(* IEC 61131-3 sources: NachHouse_TST/OSCAT_BasicLib/OscatBasicLib_333a, 28 files *)

(* ---- Arrays.ST ---- *)
TYPE
  OSCAT_BASIC_ARRAY0_32000_OF_REAL : ARRAY[0..32000] OF REAL;
  OSCAT_BASIC_ARRAY1_32000_OF_REAL : ARRAY[1..32000] OF REAL;
END_TYPE

(* @PATH := '\/Mathematical\/Array' *)
FUNCTION _ARRAY_ABS : BOOL
(*
  this function will calculate the absolute value of each element of the array and stroe the result instead of the element.
  Array[i] := ABS(ARRAY[i]).
  the function needs to be called:  array_avg(adr("array"),sizeof("array"));
  because this function works with pointers its very time efficient and it needs no extra memory.

  version 1.0 2. apr. 2008
  programmer  hugo
  tested by tobias
*)
  VAR_INPUT
    pt : PTR_TO OSCAT_BASIC_ARRAY0_32000_OF_REAL;
    size : UINT;
  END_VAR
  VAR
    i: UINT;
    stop: UINT;
  END_VAR

  stop := WORD_TO_UINT(SHR(UINT_TO_WORD(size),2))-1;
  FOR i := 0 TO stop DO
    PT^[i] := ABS(PT^[i]);
  END_FOR;
  _ARRAY_ABS := TRUE;

(* revision history
  hm  2. apr 2008   rev 1.0
    original version
*)
END_FUNCTION

(* @PATH := '\/Mathematical\/Array' *)
FUNCTION _ARRAY_ADD : BOOL
(*
  this function will add an offset X to each element of the array and stroe the result instead of the element.
  Array[i] := ARRAY[i] + X.
  the function needs to be called:  array_avg(adr("array"),sizeof("array"));
  because this function works with pointers its very time efficient and it needs no extra memory.

  version 1.0 2. apr. 2008
  programmer  hugo
  tested by tobias
*)
  VAR_INPUT
    pt : PTR_TO OSCAT_BASIC_ARRAY0_32000_OF_REAL;
    size : UINT;
    X : REAL;
  END_VAR
  VAR
    i: UINT;
    stop: UINT;
  END_VAR

  stop := WORD_TO_UINT(SHR(UINT_TO_WORD(size),2))-1; //SHR(size,2)-1;
  FOR i := 0 TO stop DO
    PT^[i] := PT^[i] + X;
  END_FOR;
  _ARRAY_ADD := TRUE;

(* revision history
  hm  2. apr 2008   rev 1.0
    original version
*)
END_FUNCTION

(* @PATH := '\/Mathematical\/Array' *)
FUNCTION _ARRAY_INIT : BOOL
(*
  this function will initialize a given array with a value init.
  the function needs to be called:  _array_init(adr("array"),sizeof("array"));
  this function will manipulate a given array.
  the function manipulates the original array, it rerturnes true when finished.
  because this function works with pointers its very time efficient and it needs no extra memory.

  version 1.3 16 mar 2008
  programmer  hugo
  tested by   tobias
*)
  VAR_INPUT
    pt : PTR_TO OSCAT_BASIC_ARRAY0_32000_OF_REAL;
    size : UINT;
    init : REAL;
  END_VAR
  VAR
    i: UINT;
    stop: UINT;
  END_VAR

  stop := WORD_TO_UINT(SHR(UINT_TO_WORD(size),2))-1; //SHR(size,2)-1;
  FOR i := 0 TO stop DO
    pt^[i] := init;
  END_FOR;

  _array_init := TRUE;

(* revision History
  hm 6.1.2007   rev 1.1
    change type of function to bool
    added  array_init := true to set output true.

  hm  14.11.2007  rev 1.2
    changed stop calculation to be more efficient

  hm  16.3. 2008    rev 1.3
    changed type of input size to uint
*)
END_FUNCTION

(* @PATH := '\/Mathematical\/Array' *)
FUNCTION _ARRAY_SORT : BOOL
(*
  this function will sort a given array.
  the function needs to be called:  _array_sort(adr("array"),sizeof("array"));
  this function will manipulate a given array.
  the function will not return anything except true, it will instead manipulate the original array.
  because this function works with pointers its very time efficient and it needs no extra memory.

  version 2.0 19. jan. 2011
  programmer  Alexander Trikitis
  tested by oscat
*)
  VAR_INPUT
    PT : PTR_TO OSCAT_BASIC_ARRAY1_32000_OF_REAL; // ARRAY[1..32000] OF REAL;
    SIZE : UINT;
  END_VAR
  VAR
    stack_count: UINT;        (* Laufvariable Stack*)
    stack: ARRAY[1..32] OF UINT;  (* Stackgröße~ 1,6*Log(n)/log(2) *)
                      (* Stackgröße 32 => ~1 Mio Elemente *)
    links: UINT;            (* Anfangselement des Arrays *)
    rechts: UINT;           (* Endelement des Arrays *)
    pivot: REAL;            (* temporärer Schwellwert für Tauschbedingung *)
    i: UINT;              (* Laufvariable1 *)
    j: UINT;              (* Laufvariable2 *)
    ende_innen: BOOL;       (* Ende innere Schleife *)
    ende_aussen: BOOL;        (* Ende äußere Schleife *)
    tmp: REAL;            (* Hilfsvariable zum Tauschen von Werten *)
  END_VAR

  (* Startwerte zur Arraygröße *)
  links := 1;         (* Anfangselement des Arrays *)
  rechts :=  WORD_TO_UINT(SHR(UINT_TO_WORD(size),2)); //SHR(size,2);    (* Endelement des Arrays *)
  stack_count := 1;     (* Laufvariable Stack *)

  WHILE NOT ende_aussen DO            (* äußere Schleife *)
    IF links < rechts THEN
      pivot := PT^[WORD_TO_UINT(SHR(UINT_TO_WORD(rechts+links),1))];      (* Wert des mittleren Elements als Pivot-Wert *)
      i := links -1;
      j := rechts +1;

      (* innere Schleife, teile Feld *)
      ende_innen := FALSE;
      REPEAT

        (* steigende Reihenfolge *)
        REPEAT  i := i+1; UNTIL (PT^[i] >= pivot) OR NOT (i < rechts) END_REPEAT;
        REPEAT  j := j-1; UNTIL (PT^[j] <= pivot) OR NOT (j > links)  END_REPEAT;

        (*sinkende Reihenfolge *)
  (*      REPEAT  i := i+1; UNTIL (PT^[i] <= pivot) OR NOT (i < rechts) END_REPEAT  *)
  (*      REPEAT  j := j-1; UNTIL (PT^[j] >= pivot) OR NOT (j > links)  END_REPEAT  *)

        IF i >= j THEN
          ende_innen := TRUE;
        ELSE
             tmp := PT^[j];
          PT^[j] := PT^[i];
          PT^[i] := tmp;
        END_IF;

      UNTIL ende_innen END_REPEAT;

      (* Push stack *)
      stack[stack_count] := rechts;   (* rechten Teil später sortieren *)
      IF Stack_count < 32 THEN
        stack_count := stack_count +1;
      ELSE
        ende_aussen := TRUE;
        _ARRAY_SORT := FALSE;         (* Fehler: Stack zu klein *)
      END_IF;

      (* linken Teil sortiern *)
      rechts := MAX(links, i-1);

    ELSE

      IF stack_count = 1 THEN
        ende_aussen := TRUE;
      ELSE

        links := rechts+1;

        (* pop stack *)
        stack_count := stack_count -1;    (* jetzt rechten Teil sortierne *)
        rechts:= stack[stack_count];
      END_IF;

    END_IF;

  END_WHILE;

  _ARRAY_SORT := TRUE;        (* Sortierung beendet *)

(* algorithm used before rev 2.0
  size := SHR(size,2);
  size2 := UINT_TO_INT(SHR(size,1));
  FOR i := SIZE2  TO 1 BY -1 DO
    j:=i;
      WHILE j <= SIZE2 DO
        stop := j * 2 + 1;
          IF stop > UINT_TO_INT(SIZE) THEN stop := stop - 1;
          ELSIF pt^[stop-1] > pt^[stop] THEN stop := stop - 1;
      END_IF;
          IF pt^[j] < pt^[stop] THEN
            temp := pt^[j];
              pt^[j] := pt^[stop];
              pt^[stop] := temp;
          END_IF;
          j := stop;
      END_WHILE;
  END_FOR;
*)

(* heapsort
  FOR heapsize := UINT_TO_INT(size) TO 1 BY -1 DO
    popmax := pt^[1];
    pt^[1] := pt^[heapsize];
      i := 1;
    hs2 := SHR(heapsize,1);
    WHILE i <= hs2 DO
          stop := i * 2 + 1;
            IF stop > heapsize THEN stop := stop - 1;
            ELSIF pt^[stop-1] > pt^[stop] THEN stop := stop - 1;
      END_IF;
            IF pt^[i] < pt^[stop] THEN
                  temp := pt^[i];
                  pt^[i] := pt^[stop];
                  pt^[stop] := temp;
            END_IF;
            i := stop;
        END_WHILE;
    pt^[heapsize] := popmax;
  END_FOR;

  _ARRAY_SORT2 := TRUE;
*)

(* old algorithm bubble sort used before rev 1.2
  stop := (size - SIZEOF(pt)) / SIZEOF(pt);
  FOR i := 0 TO stop - 1 DO
    FOR m := i + 1 TO stop DO
      IF pt^[i] > pt^[m] THEN
        temp := pt^[i];
        pt^[i] := pt^[m];
        pt^[m] := temp;
      END_IF;
    END_FOR;
  END_FOR;
  _array_sort := TRUE;
*)

(* revision history
  hm  6.1.2007  rev 1.1
    changed return value to true

  hm  22. sep 2007  rev 1.2
    changed sorting algorithm to heap sort for performance reasons

  hm  14. nov 2007  rev 1.3
    changed calculation of stop to be more efficient

  hm  15 dec 2007 rev 1.4
    added function return true

  hm  5. jan 2008   rev 1.5
    improved performance

  hm  16. mar. 2008 rev 1.6
    changed type of input size to uint

  hm  28. mar. 2008 rev 1.7
    changed input f to pt

  hm  19. jan. 2011 rev 2.0
    new faster algorithm using qucksort (Alexander Drikitis)
*)
END_FUNCTION

(* @PATH := '\/Mathematical\/Array' *)
FUNCTION _ARRAY_MEDIAN : REAL
(*
  this function will calculate the median of a given array.
  in order to do so the ariginal array is sorted and stays sorted after the function finishes
  the function needs to be called:  _array_median(adr("array"),sizeof("array"));
  this function will manipulate a given array.
  the function will return the median of the original array.
  for example [12,0,4,7,1] the median is 4 and the array after the function is called is [0,1,4,7,12]
  because this function works with pointers its very time efficient and it needs no extra memory.

  version 1.5 16 mar 2008
  programmer  hugo
  tested by   tobias
*)
  VAR_INPUT
    pt : PTR_TO OSCAT_BASIC_ARRAY0_32000_OF_REAL;
    size : UINT;
  END_VAR
  VAR
    i: UINT;
    stop: UINT;
  END_VAR

  _ARRAY_SORT(pt,size);
  stop := WORD_TO_UINT(SHR(UINT_TO_WORD(size),2))-1; //SHR(size,2)-1;
  IF EVEN(UINT_TO_DINT(stop)) THEN
    _ARRAY_MEDIAN := pt^[WORD_TO_UINT(SHR(UINT_TO_WORD(stop),1))];
  ELSE
    i := WORD_TO_UINT(SHR(UINT_TO_WORD(stop),1));
    _ARRAY_MEDIAN := (pt^[i] + pt^[i+1]) * 0.5;
  END_IF;

(* old code
  stop := (size - SIZEOF(pt)) / SIZEOF(pt);
  FOR i := 0 TO stop - 1 DO
    FOR m := i + 1 TO stop DO
      IF pt^[i] > pt^[m] THEN
        temp := pt^[i];
        pt^[i] := pt^[m];
        pt^[m] := temp;
      END_IF;
    END_FOR;
  END_FOR;
  IF even(stop) THEN
    _array_median := pt^[stop/2];
  ELSE
    i := stop/2;
    _array_median := (pt^[i] + pt^[i+1])/2;
  END_IF;
*)
(* revision history
  hm  3.3.2007    rev 1.1
    corrected an error, changed the statement line 14 i := TRUNC(stop/2); to i := stop/2;

  hm    22. sep 2007  rev 1.2
    changed algorithm to use _array_soft for performance reasons

  hm    8. oct 2007   rev 1.3
    deleted unused variables m and temp

  hm    14. nov 2007  rev 1.4
    corrected a problem with size calculation

  hm    16.3. 2008    rev 1.5
    changed type of input size to uint
    performance improvements
*)
END_FUNCTION

(* @PATH := '\/Mathematical\/Array' *)
FUNCTION _ARRAY_MUL : BOOL
(*
  this function will multiply each element of the array and stroe the result instead of the element.
  Array[i] := ARRAY[i] * X.
  the function needs to be called:  array_avg(adr("array"),sizeof("array"));
  because this function works with pointers its very time efficient and it needs no extra memory.

  version 1.0 2. apr. 2008
  programmer  hugo
  tested by tobias
*)
  VAR_INPUT
    pt : PTR_TO OSCAT_BASIC_ARRAY0_32000_OF_REAL;
    size : UINT;
    X : REAL;
  END_VAR
  VAR
    i: UINT;
    stop: UINT;
  END_VAR

  stop := WORD_TO_UINT(SHR(UINT_TO_WORD(size),2))-1; //SHR(size,2)-1;
  FOR i := 0 TO stop DO
    PT^[i] := PT^[i] * X;
  END_FOR;
  _ARRAY_MUL := TRUE;

(* revision history
  hm  2. apr 2008   rev 1.0
    original version
*)
END_FUNCTION

(* @PATH := '\/Mathematical\/Array' *)
FUNCTION _ARRAY_SHUFFLE : BOOL
(*
  this function will randomly shuffle the elements of an array

  version 1.2 30. mar. 2008
  programmer  kurt
  tested by   hugo
*)
  VAR_INPUT
    pt : PTR_TO OSCAT_BASIC_ARRAY0_32000_OF_REAL;
    size : UINT;
  END_VAR
  VAR
    temp : REAL;
    pos  : INT;
    i: INT;
    stop: INT;
  END_VAR

  stop := WORD_TO_INT(SHR(UINT_TO_WORD(size),2))-1; //UINT_TO_INT(SHR(size,2)-1);
  FOR i := 0 TO stop DO
          pos := RDM2(i+pos,0,stop);
          (* swap elements *)
          temp := pt^[i];
          pt^[i] := pt^[pos];
          pt^[pos] := temp;
  END_FOR;

  _ARRAY_SHUFFLE := TRUE;

(* revision History
  hm  4. mar 2008 rev 1.0
    original version

  hm  16. mar. 2008 rev 1.1
    changed type of input size to uint

  hm  30. mar. 2008 rev 1.2
    changed last in rdm2 fromm pos to i + pos to allow for more randomness
*)
END_FUNCTION

(* @PATH := '\/Mathematical\/Array' *)
FUNCTION ARRAY_AVG : REAL
(*
  this function will calculate the average of a given array.
  the function needs to be called:  array_avg(adr("array"),sizeof("array"));
  because this function works with pointers its very time efficient and it needs no extra memory.

  version 1.3 10. mar. 2009
  programmer  hugo
  tested by   tobias
*)
  VAR_INPUT
    pt : PTR_TO OSCAT_BASIC_ARRAY0_32000_OF_REAL;
    size : UINT;
  END_VAR
  VAR
    i: UINT;
    stop: UINT;
  END_VAR
  VAR_TEMP
    tmp : REAL;
  END_VAR

  stop := WORD_TO_UINT(SHR(UINT_TO_WORD(size),2))-1; //SHR(size,2)-1;
  tmp := pt^[0];
  FOR i := 1 TO stop DO
    tmp := tmp + pt^[i];
  END_FOR;
  tmp := tmp / UINT_TO_REAL(stop + 1);
  ARRAY_AVG := tmp;

(* revision history
  hm  2. oct 2007   rev 1.0
    original version

  hm  12. dec 2007  rev 1.1
    chaged code for better performance

  hm  16. mar. 2008 rev 1.2
    changed input size to uint

  hm  10. mar. 2009 rev 1.3
    added type conversion for compatibility reasons
*)
END_FUNCTION

(* @PATH := '\/Mathematical\/Array' *)
FUNCTION ARRAY_GAV : REAL
(*
  this function will calculate the geometric average of a given array.
  the function needs to be called:  array_avg(adr("array"),sizeof("array"));
  because this function works with pointers its very time efficient and it needs no extra memory.

  version 1.1 10. mar. 2009
  programmer  hugo
  tested by   tobias
*)
  VAR_INPUT
    pt : PTR_TO OSCAT_BASIC_ARRAY0_32000_OF_REAL;
    size : UINT;
  END_VAR
  VAR
    i: UINT;
    stop: UINT;
  END_VAR
  VAR_TEMP
    tmp : REAL;
  END_VAR

  stop := WORD_TO_UINT(SHR(UINT_TO_WORD(size),2))-1; //SHR(size,2)-1;
  tmp := 1.0;
  FOR i := 0 TO stop DO
    IF pt^[i] > 0.0 THEN
      tmp := tmp * pt^[i];
    ELSE
      tmp := 0.0;
      RETURN;
    END_IF;
  END_FOR;
  tmp := SQRTN(tmp,UINT_TO_INT(stop)+1);
  ARRAY_GAV := tmp;

(* revision history
  hm  2. apr 2008 rev 1.0
    original version

  hm  10. mar. 2009 rev 1.1
    real constants updated to new systax using dot
*)
END_FUNCTION

(* @PATH := '\/Mathematical\/Array' *)
FUNCTION ARRAY_HAV : REAL
(*
  this function will calculate the harmonic average of a given array.
  the function needs to be called:  array_avg(adr("array"),sizeof("array"));
  because this function works with pointers its very time efficient and it needs no extra memory.

  version 1.1 10. mar. 2009
  programmer  hugo
  tested by   tobias
*)
  VAR_INPUT
    pt : PTR_TO OSCAT_BASIC_ARRAY0_32000_OF_REAL;
    size : UINT;
  END_VAR
  VAR
    i: UINT;
    stop: UINT;
  END_VAR
  VAR_TEMP
    tmp : REAL;
  END_VAR

  stop := WORD_TO_UINT(SHR(UINT_TO_WORD(size),2))-1; //SHR(size,2)-1;
  FOR i := 0 TO stop DO
    IF pt^[i] <> 0.0 THEN
      tmp := tmp + 1.0 / pt^[i];
    ELSE
      tmp := 0.0;
      RETURN;
    END_IF;
  END_FOR;
  tmp := UINT_TO_REAL(stop + 1) / tmp;
  ARRAY_HAV := tmp;

(* revision history
  hm  2. apr 2008 rev 1.0
    original version

  hm  10. mar. 2009 rev 1.1
    real constants updated to new systax using dot
*)
END_FUNCTION

(* @PATH := '\/Mathematical\/Array' *)
FUNCTION ARRAY_MAX : REAL
(*
  this function will calculate the max value of a given array.
  the function needs to be called:  array_max(adr("array"),sizeof("array"));
  because this function works with pointers its very time efficient and it needs no extra memory.

  version 1.1 16. mar. 2008
  programmer  hugo
  tested by   tobias
*)
  VAR_INPUT
    pt : PTR_TO OSCAT_BASIC_ARRAY0_32000_OF_REAL;
    size : UINT;
  END_VAR
  VAR
    i: UINT;
    stop: UINT;
  END_VAR
  VAR_TEMP
    tmp : REAL;
  END_VAR

  stop := (size -SIZEOF(pt)) / SIZEOF(pt);
  tmp := pt^[0];
  FOR i := 1 TO stop DO
    IF pt^[i] > tmp THEN tmp := pt^[i]; END_IF;
  END_FOR;
  ARRAY_MAX := tmp;

(* revision history
  hm  2. oct 2006   rev 1.0
    original version

  hm  16. mar. 2008 rev 1.1
    changed input size to uint
*)
END_FUNCTION

(* @PATH := '\/Mathematical\/Array' *)
FUNCTION ARRAY_MIN : REAL
(*
  this function will calculate the min value of a given array.
  the function needs to be called:  array_min(adr("array"),sizeof("array"));
  because this function works with pointers its very time efficient and it needs no extra memory.

  version 1.1 16. mar. 2008
  programmer  hugo
  tested by   tobias
*)
  VAR_INPUT
    pt : PTR_TO OSCAT_BASIC_ARRAY0_32000_OF_REAL;
    size : UINT;
  END_VAR
  VAR
    i: UINT;
    stop: UINT;
  END_VAR
  VAR_TEMP
    tmp : REAL;
  END_VAR

  stop := (size - SIZEOF(pt)) / SIZEOF(pt);
  tmp := pt^[0];
  FOR i := 1 TO stop DO
    IF pt^[i] < tmp THEN tmp := pt^[i]; END_IF;
  END_FOR;
  ARRAY_MIN := tmp;

(* revision history
  hm    2. oct. 2006
    original version

  hm    16. mar. 2008
    changed type of input size to uint
*)
END_FUNCTION

(* @PATH := '\/Mathematical\/Array' *)
FUNCTION ARRAY_VAR : REAL
(*
  this function will calculate the variance of a given array.
  the function needs to be called:  array_var(adr("array"),sizeof("array"));
  because this function works with pointers its very time efficient and it needs no extra memory.

  version 1.3 10. mar. 2009
  programmer  hugo
  tested by   tobias
*)
  VAR_INPUT
    pt : PTR_TO OSCAT_BASIC_ARRAY0_32000_OF_REAL;
    size : UINT;
  END_VAR
  VAR
    avg : REAL;
    i: UINT;
    stop: UINT;
  END_VAR
  VAR_TEMP
    tmp : REAL;
  END_VAR

  (* at first we calualte the arithmetic average of the array *)

  stop := WORD_TO_UINT(SHR(UINT_TO_WORD(size),2))-1; //SHR(size,2)-1;
  avg := pt^[0];
  FOR i := 1 TO stop DO
    avg := avg + pt^[i];
  END_FOR;
  avg := avg / UINT_TO_REAL(stop + 1);

  (* in a second run we calculate the variance of the array *)

  tmp := (pt^[0] - avg) * (pt^[0] - avg);
  FOR i := 1 TO stop DO
    tmp := tmp + (pt^[i] - avg) * (pt^[i] - avg);
  END_FOR;
  ARRAY_VAR := tmp / UINT_TO_REAL(stop);

(* revision history
  hm  1.4.2007  rev 1.0
    function created

  hm  12.12.2007  rev 1.1
    changed code for better performance

  hm  16. mar. 2008 rev 1.2
    changed type of input size to uint

  hm  10. mar. 2009 rev 1.3
    added type conversions for compatibility reasons
*)
END_FUNCTION

(* @PATH := '\/Mathematical\/Array' *)
FUNCTION ARRAY_SDV : REAL
(*
  this function will calculate the standard deviation of a given array.
  the function needs to be called:  array_sdv(adr("array"),sizeof("array"));
  because this function works with pointers its very time efficient and it needs no extra memory.

  version 1.1 16. mar 2008
  programmer  hugo
  tested by   tobias
*)
  VAR_INPUT
    pt : PTR_TO OSCAT_BASIC_ARRAY0_32000_OF_REAL;
    size : UINT;
  END_VAR

  (* standard deviation is simply the square root of the variance *)
  array_sdv := SQRT( array_var(pt, size));

(* revision history
  hm  1.4.2007    rev 1.0
    function created

  hm  16. mar. 2008 rev 1.1
    changed type of input size to uint
*)
END_FUNCTION

(* @PATH := '\/Mathematical\/Array' *)
FUNCTION ARRAY_SPR : REAL
(*
  this function will calculate the spread of a given array.
  the function needs to be called:  array_spr(adr("array"),sizeof("array"));
  for example: spread of [12,0,4,1,7] is 12 - 0 = 12.
  because this function works with pointers its very time efficient and it needs no extra memory.

  version 1.1 16. mar. 2008
  programmer  hugo
  tested by   tobias
*)
  VAR_INPUT
    pt : PTR_TO OSCAT_BASIC_ARRAY0_32000_OF_REAL;
    size : UINT;
  END_VAR
  VAR
    i: UINT;
    stop: UINT;
    array_max : REAL;
    array_min : REAL;
  END_VAR

  stop := (size -SIZEOF(pt)) / SIZEOF(pt);
  array_min := pt^[0];
  array_max := pt^[0];
  FOR i := 1 TO stop DO
    IF pt^[i] > array_max THEN array_max := pt^[i];
    ELSIF pt^[i] < array_min THEN array_min := pt^[i];
    END_IF;
  END_FOR;
  array_spr := array_max - array_min;

(* revision history
  hm  2. oct. 2006  rev 1.0
    original version

  hm  16. mar. 2008 rev 1.1
    changed type of input size to uint
*)
END_FUNCTION

(* @PATH := '\/Mathematical\/Array' *)
FUNCTION ARRAY_SUM : REAL
(*
  this function will calculate the sum of a given array.
  the function needs to be called:  array_sum(adr("array"),sizeof("array"));
  because this function works with pointers its very time efficient and it needs no extra memory.

  version 1.1 16. mar. 2008
  programmer  hugo
  tested by   tobias
*)
  VAR_INPUT
    pt : PTR_TO OSCAT_BASIC_ARRAY0_32000_OF_REAL;
    size : UINT;
  END_VAR
  VAR
    i: UINT;
    stop: UINT;
  END_VAR
  VAR_TEMP
    tmp : REAL;
  END_VAR

  stop := (size -SIZEOF(pt)) / SIZEOF(pt);
  tmp := pt^[0];
  FOR i := 1 TO stop DO
    tmp := tmp + pt^[i];
  END_FOR;
  ARRAY_SUM := tmp;

(* revision history
  hm  2. oct. 2006  rev 1.0
    function created

  hm  16. mar. 2008 rev 1.1
    changed type of input size to uint
*)
END_FUNCTION

(* @PATH := '\/Mathematical\/Array' *)
FUNCTION ARRAY_TREND : REAL
(*
  this function will calculate the trend of a given array.
  trend will calculate the avg of the first half of the array and then the avg of the second half, trend = avg2 - avg1.
  for example:  [0,1,4,5,3,4,6,3] = 4 - 2.5 = 1.5
  the function needs to be called:  array_trend(adr("array"),sizeof("array"));
  because this function works with pointers its very time efficient and it needs no extra memory.

  version 1.3 10. mar. 2009
  programmer  hugo
  tested by   tobias
*)
  VAR_INPUT
    pt : PTR_TO OSCAT_BASIC_ARRAY0_32000_OF_REAL;
    size : UINT;
  END_VAR
  VAR
    i: UINT;
    stop: UINT;
    x: REAL;
    stop2: UINT;
  END_VAR

  stop := WORD_TO_UINT(SHR(UINT_TO_WORD(size),2))-1; //SHR(size,2)-1;
  stop2 := WORD_TO_UINT(SHR(UINT_TO_WORD(stop),1));  //SHR(stop,1);
  FOR i := 0 TO stop2 DO x := x - pt^[i]; END_FOR;
  IF EVEN(UINT_TO_DINT(stop)) THEN
    FOR i := stop2 TO stop DO X := X + pt^[i]; END_FOR;
  ELSE
    FOR i := stop2 + 1 TO stop DO X := X + pt^[i]; END_FOR;
  END_IF;
  ARRAY_TREND := x / UINT_TO_REAL(stop2 + 1);

(* revision history
  hm  2 oct 2007  rev 1.0
    original version

  hm  12 dec 2007 rev 1.1
    changed code for better performance

  hm  16. mar. 2008 rev 1.2
    changed type of input size to uint

  hm  10. mar. 2009 rev 1.3
    added type conversions for compatibility reasons
*)
END_FUNCTION

(* @PATH := '\/Mathematical\/Array' *)
FUNCTION IS_SORTED : BOOL
(*
  this function will return true if the given array is sorted in an ascending order.
  the function needs to be called:  array_sorted(adr("array"),sizeof("array"));
  because this function works with pointers its very time efficient and it needs no extra memory.

  version 1.1 4. apr. 2008
  programmer  hugo
  tested by tobias
*)
  VAR_INPUT
    pt : PTR_TO OSCAT_BASIC_ARRAY0_32000_OF_REAL;
    size : UINT;
  END_VAR
  VAR
    stop: INT;
    i: INT;
  END_VAR

  stop := WORD_TO_INT(SHR(UINT_TO_WORD(size),2))-2; //UINT_TO_INT(SHR(size,2)-2);
  FOR i := 0 TO stop DO
    IF pt^[i] > pt^[i+1] THEN
      IS_SORTED := FALSE;
      RETURN;
    END_IF;
  END_FOR;

  IS_SORTED := TRUE;

(* revision history
  hm  29. mar. 2008   rev 1.0
    original version

  hm  4. apr. 2008  rev 1.1
    added type conversion to avoid warnings under codesys 3.0
*)
END_FUNCTION

(* ---- BUFFER_Management.ST ---- *)
TYPE
  OSCAT_BASIC_ARRAY0_32767_OF_BYTE : ARRAY[0..32767] OF BYTE;
  OSCAT_BASIC_ARRAY0_STRING_LENGTH_OF_BYTE : ARRAY[0..STRING_LENGTH] OF BYTE;
END_TYPE

(* @PATH := '\/Buffer Management' *)
FUNCTION _BUFFER_CLEAR : BOOL
(*
  this function will initialize a given array of byte with 0.
  the function needs to be called:	_buffer_clear(adr("array"),sizeof("array"));
  this function will manipulate a given array.
  the function manipulates the original array, it rerturnes true when finished.
  because this function works with pointers its very time efficient and it needs no extra memory.

  version 1.2	31. oct. 2008
  programmer 	hugo
  tested by	oscat
*)
  VAR_INPUT
  	PT : PTR_TO BYTE;
  	SIZE : UINT;
  END_VAR
  VAR
  	ptw        : PTR_TO DWORD;
  	temp       : UDINT;
  	end, end32 : UDINT;
  END_VAR

  (* this routine uses 32 bit access to gain speed *)
  (* first access bytes till pointer is aligned for 32 bit access *)
  temp := PTR_TO_UDINT( pt);
  end := temp + UINT_TO_UDINT(size);
  end32 := end - 3;
  WHILE (PTR_TO_UDINT(pt) < end) AND ((UDINT_TO_DWORD(temp) AND 16#00000003) > 0) DO
  	pt^ := 0;
  	pt := pt + 1;
  	temp := temp + 1;
  END_WHILE;
  (* pointer is aligned, now copy 32 bits at a time *)
  ptw := pt;
  WHILE PTR_TO_UDINT(ptw) < end32 DO (* *)
  	ptw^ := 0;
  	ptw := ptw + 4;
  END_WHILE;
  (* copy the remaining bytes in byte mode *)
  pt := ptw;
  WHILE PTR_TO_UDINT(pt) < end DO
  	pt^ := 0;
  	pt := pt + 1;
  END_WHILE;
  _BUFFER_CLEAR := TRUE;

(* revision History
  hm 	5. mar. 2008	rev 1.0
  	original version

  hm	16. mar. 2008	rev 1.1
  	added type conversion to avoid warnings under codesys 30
  	chaged type of input size to uint
  	deleted unused variable i

  hm	31. oct. 2008	rev 1.2
  	corrected an error while routine would write outside of arrays
  *)
END_FUNCTION

(* @PATH := '\/Buffer Management' *)
FUNCTION _BUFFER_INIT : BOOL
(*
  this function will initialize a given array of byte with init.
  the function needs to be called:	_buffer_init(adr("array"),sizeof("array"),init);
  this function will manipulate a given array.
  the function manipulates the original array, it rerturnes true when finished.
  because this function works with pointers its very time efficient and it needs no extra memory.

  version 1.2	31. oct. 2008
  programmer 	hugo
  tested by	oscat
*)
  VAR_INPUT
  	PT : PTR_TO BYTE;
  	SIZE : UINT;
  	INIT : BYTE;
  END_VAR
  VAR
  	ptw : PTR_TO UDINT;
  	temp : UDINT;
  	end, end32 : UDINT;
  END_VAR

  (* this routine uses 32 bit access to gain speed *)
  (* first access bytes till pointer is aligned for 32 bit access *)
  temp := PTR_TO_UDINT(pt);
  end := temp + UINT_TO_UDINT(size);
  end32 := end - 3;
  WHILE (PTR_TO_UDINT(pt) < end) AND ((UDINT_TO_DWORD(temp) AND 16#00000003) > 0) DO
  	pt^ := init;
  	pt := pt + 1;
  	temp := temp + 1;
  END_WHILE;
  (* pointer is aligned, now copy 32 bits at a time *)
  ptw := pt;
  temp := DWORD_TO_UDINT( SHL(BYTE_TO_DWORD(init),24) OR SHL(BYTE_TO_DWORD(init),16) OR SHL(BYTE_TO_DWORD(init),8) OR BYTE_TO_DWORD(init));
  WHILE PTR_TO_UDINT(ptw) < end32 DO
  	ptw^ := temp;
  	ptw := ptw + 4;
  END_WHILE;
  (* copy the remaining bytes in byte mode *)
  pt := ptw;
  WHILE PTR_TO_UDINT(pt) < end DO
  	pt^ := init;
  	pt := pt + 1;
  END_WHILE;
  _BUFFER_INIT := TRUE;

(* revision History
  hm 	5. mar. 2008	rev 1.0
  	original version

  hm	16. mar. 2008	rev 1.1
  	added type conversion to avoid warnings under codesys 3.0
  	chaged type of input size to uint.

  hm	31. oct. 2008	rev 1.2
  	corrected an error while routine would write outside of arrays
  *)
END_FUNCTION

(* @PATH := '\/Buffer Management' *)
FUNCTION _STRING_TO_BUFFER : INT
(*
  this function will copy a string into an array of byte starting at position pos.
  the function needs to be called:	_String_To_buffer(str, pos, adr("array"),sizeof("array"));
  this function will manipulate the array directly in memory and returns the position after the input string when finished.
  because this function works with pointers its very time efficient and it needs no extra memory.

  version 1.4	2. jan. 2012
  programmer 	hugo
  tested by		oscat
*)
  VAR_INPUT
  	STR : STRING[STRING_LENGTH];
  	POS : INT;
  	PT : PTR_TO OSCAT_BASIC_ARRAY0_32767_OF_BYTE; // ARRAY[0..32767] OF BYTE;
  	SIZE : UINT;
  END_VAR
  VAR
  	ps : PTR_TO BYTE;
  	i: INT;
  	end: INT;
  END_VAR

  ps := ADR(str);
  end := MIN(pos + LEN(str), UINT_TO_INT(size));
  IF end > 0 THEN end := end -1; END_IF;
  FOR i := pos TO end DO
  	pt^[i] := ps^;
  	ps := ps + 1;
  END_FOR;
  _STRING_TO_BUFFER := i;

(* revision History

  hm 	5. mar. 2008	rev 1.0
  	original version

  hm	16. mar. 2008	rev 1.1
  	changed type of input size to uint

  hm	13. may. 2008	rev 1.2
  	changed type of pointer to array[1..32767]
  	changed size of string to STRING_LENGTH

  hm	12. nov. 2009	rev 1.3
  	limit end to size - 1

  hm	2. jan 2012	rev 1.4
  	return the position after the input string when finished
*)
END_FUNCTION

(* @PATH := '\/Buffer Management' *)
FUNCTION _BUFFER_INSERT : INT
(*
  this function will insert a string at a given position in a buffer.
  the function needs to be called:	_buffer_insert(str, pos, adr("array"), sizeof("array"));
  this function will manipulate a given array.
  the function manipulates the original array, it returnes the next position after the input string when finished.
  because this function works with pointers its very time efficient and it needs no extra memory.

  version 1.5	2. jan. 2012
  programmer 	hugo
  tested by	oscat
*)
  VAR_INPUT
  	STR : STRING[STRING_LENGTH];
  	POS : INT;
  	PT : PTR_TO OSCAT_BASIC_ARRAY0_32767_OF_BYTE; // ARRAY[0..32767] OF BYTE;
  	SIZE : UINT;
  END_VAR
  VAR
  	end : INT;
  	lx: INT;
  	i: INT;
  END_VAR

  lx := LEN(str);
  end := pos + lx;
  (* first move the upper part of the buffer to make space for the string *)
  FOR i := UINT_TO_INT(size) - 1 TO end BY -1 DO
  	pt^[i] := pt^[i-lx];
  END_FOR;
  (* copy the string *)
  _BUFFER_INSERT := _STRING_TO_BUFFER(str, pos, PT, size);

(* revision History
  hm 	9. mar. 2008	rev 1.0
  	original version

  hm	16. mar. 2008	rev 1.1
  	changed type of input size to uint

  hm	13. may. 2008	rev 1.2
  	changed type of pointer to array[1..32767]
  	changed size of string to STRING_LENGTH

  hm	23. mar. 2009	rev 1.3
  	avoid writing to input pos

  hm	12. nov. 2009	rev 1.4
  	code optimized

  hm 2. jan 2012	rev 1.5
  	function now returns the next position after the input string
*)
END_FUNCTION

(* @PATH := '\/Buffer Management' *)
FUNCTION _BUFFER_UPPERCASE : BOOL
(*
  this function will convert an array of byte into uppercase
  the function needs to be called:  _buffer_clear(adr("array"),sizeof("array"));
  this function will manipulate a given array.
  the function manipulates the original array, it rerturnes true when finished.
  because this function works with pointers its very time efficient and it needs no extra memory.

  version 1.0 20. jan. 2011
  programmer  hugo
  tested by oscat
*)
  VAR_INPUT
    PT : PTR_TO OSCAT_BASIC_ARRAY0_32767_OF_BYTE; //ARRAY[0..32000] OF BYTE;
    SIZE : INT;
  END_VAR
  VAR
    pos: INT;
  END_VAR

  pos := 0;
  WHILE pos < size DO
    PT^[pos] := TO_UPPER(pt^[pos]);
    pos := pos + 1;
  END_WHILE;
  _BUFFER_UPPERCASE := TRUE;

(* revision History
  hm  20. jan. 2011 rev 1.0
    original version
*)
END_FUNCTION

(* @PATH := '\/Buffer Management' *)
FUNCTION BUFFER_COMP : INT
(*
  version 1.1 12. nov. 2009
  programmer  hugo
  tested by oscat
*)
  VAR_INPUT
    PT1 : PTR_TO OSCAT_BASIC_ARRAY0_32767_OF_BYTE; // ARRAY[0..32767] OF BYTE;
    SIZE1 : INT;
    PT2 : PTR_TO OSCAT_BASIC_ARRAY0_32767_OF_BYTE; // ARRAY[0..32767] OF BYTE;
    SIZE2 : INT;
    START : INT;
  END_VAR
  VAR
    i, j, end : INT;
    firstbyte: BYTE;
  END_VAR

  (* search for first character match *)
  IF size2 <= size1 THEN
    end := size1 - size2;
    firstbyte := PT2^[0];
    FOR i := START TO end DO
      IF PT1^[i] = firstbyte THEN
        (* first character matches, now compare rest of array *)
        j := 1;
        WHILE j < size2 DO
          IF pt2^[j] <> pt1^[j+i] THEN EXIT; END_IF;
          j := j + 1;
        END_WHILE;
        (* when J > size2 a match was found return the position i in buffer1 *)
        IF j = size2 THEN
          BUFFER_COMP := i;
          RETURN;
        END_IF;
      END_IF;
    END_FOR;
  END_IF;
  BUFFER_COMP := -1;

(*
  hm 14. nov. 2008  rev 1.0
    original version

  hm  12. nov. 2009 rev 1.1
    performance increase
*)
END_FUNCTION

(* @PATH := '\/Buffer Management' *)
FUNCTION BUFFER_SEARCH : INT
(*
  this function will search for a string STR in an array of byte starting at position pos.
  the function needs to be called: buffer_search(adr("array"),sizeof("array"), STR, POS, IGN);
  because this function works with pointers its very time efficient and it needs no extra memory.
  The function returns the position of the first character of the string in the array if found.
  a -1 is returned if the string is not found in the array.
  when IGN = TRUE, STR must be in capital letters and the search is case insensitv.

  version 1.4 25. jan 2011
  programmer  hugo
  tested by oscat
*)
  VAR_INPUT
    PT : PTR_TO OSCAT_BASIC_ARRAY0_32767_OF_BYTE; // ARRAY[0..32767] OF BYTE;
    SIZE : INT;
    STR : STRING[STRING_LENGTH];
    POS : INT;
    IGN : BOOL;
  END_VAR
  VAR
    ps : PTR_TO OSCAT_BASIC_ARRAY0_STRING_LENGTH_OF_BYTE; // ARRAY[0..STRING_LENGTH] OF BYTE;
    chx : BYTE;
    i: INT;
    end: INT;
    k: INT;
    lx: INT;
  END_VAR

  ps := ADR(STR);
  lx := LEN(STR);
  end := MIN(SIZE - lx, SIZE - 1);
  lx := lx - 1;
  FOR i := pos TO end DO
    FOR k := 0 TO lx DO
      IF IGN THEN chx := TO_UPPER(pt^[i+k]); ELSE chx := pt^[i+k]; END_IF;
      IF ps^[k] <> chx THEN EXIT; END_IF;
    END_FOR;
    IF k > lx THEN
      BUFFER_SEARCH := i;
      RETURN;
    END_IF;
  END_FOR;
  BUFFER_SEARCH := -1;

(* revision History
  hm 5. mar. 2008 rev 1.0
    original version

  hm  16. mar. 2008 rev 1.1
    chaged type of input size to uint

  hm  13. may. 2008 rev 1.2
    changed type of pointer to array[1..32767]
    changed size of string to STRING_LENGTH

  hm  12. nov. 2009 rev 1.3
    limit end to array size

  hm  25. jan. 2011 rev 1.4
    ign = True will now ignore case
    return -1 if nothing found
*)
END_FUNCTION

(* @PATH := '\/Buffer Management' *)
FUNCTION BUFFER_TO_STRING : STRING[STRING_LENGTH]
(*
  this function will retrieve a string from an array of byte starting at position start and stop at position stop.
  the function needs to be called:  buffer_TO_String(adr("array"),sizeof("array"), start, stop);
  because this function works with pointers its very time efficient and it needs no extra memory.

  version 1.5 12. nov. 2009
  programmer  hugo
  tested by   oscat
*)
  VAR_INPUT
    PT : PTR_TO OSCAT_BASIC_ARRAY0_32767_OF_BYTE; // ARRAY[0..32767] OF BYTE;
    SIZE : UINT;
    START : UINT;
    STOP : UINT;
  END_VAR
  VAR
    ps : PTR_TO BYTE;
    i : UINT;
    stp: UINT;
    sta: UINT;
  END_VAR

  ps := ADR(BUFFER_TO_STRING);
  IF size = 0 THEN RETURN; END_IF;
  sta := MIN(start, size -1);
  stp := MIN(stop, size -1);

  (* check for maximum string_length *)
  IF UINT_TO_INT(stp - sta + 1) >= STRING_LENGTH THEN
    stp := sta + INT_TO_UINT(STRING_LENGTH) - 1;
  END_IF;

  FOR i := sta TO stp DO
    ps^ := pt^[i];
    ps := ps + 1;
  END_FOR;

  (* terminate the string *)
  ps^ := 0;

(* revision History
  hm  5. mar. 2008  rev 1.0
    original version

  hm  16. mar. 2008 rev 1.1
    changed type of input size to uint

  hm  13. may. 2008 rev 1.2
    changed type of pointer to array[0..32767]
    changed size of string to STRING_LENGTH

  hm  12. jun. 2008 rev 1.3
    check for pointer overrun
    change input start and stop to uint
    added type conversions to avoid warnings under codesys 3.0

  hm  23. mar. 2009 rev 1.4
    avoid writing to input stop

  hm  12. nov. 2009 rev 1.5
    limit start and stop to size -1
*)
END_FUNCTION

(* ---- List_Processing.ST ---- *)
TYPE
  OSCAT_BASIC_ARRAY1_LIST_LENGTH_OF_BYTE : ARRAY[1..LIST_LENGTH] OF BYTE;
END_TYPE

(* @PATH := '\/List Processing' *)
FUNCTION LIST_ADD : BOOL
(*
  LIST_ADD hängt ein weiteres element ans ende einer liste.
  die liste liegt als string von elementen vor die mit den zeichen SEP am anfang makiert sind.

  version 2.0   21. mar. 2011
  programmer  hugo
  tested by   kurt
*)
  VAR_INPUT
    SEP : BYTE;
    INS : STRING[LIST_LENGTH];
  END_VAR
  VAR_IN_OUT
    LIST : STRING[LIST_LENGTH];
  END_VAR
  VAR
    sx : STRING[1];
  END_VAR

  sx := CHR_TO_STRING(SEP);     (* convert separation character to string *)
  INS := CONCAT(sx, INS);         (* start element with separation character *)

  IF LEN(LIST) + LEN(INS) > LIST_LENGTH THEN
    LIST_ADD := FALSE;          (* return false if element does not fit *)
  ELSE
    LIST := CONCAT(LIST, INS);
    LIST_ADD := TRUE;
  END_IF;

(* revision histroy
  hm  21. mar. 2011 rev 2.0
    original release
*)
END_FUNCTION

(* @PATH := '\/List Processing' *)
FUNCTION LIST_CLEAN : BOOL
(*
  LIST_CLEAN bereinigt eine liste von leeren Elementen.
  die liste liegt als string von elementen vor die mit den zeichen SEP am anfang markiert sind.

  version 2.0 21. mar. 2011
  programmer  hugo
  tested by   oscat
*)
  VAR_INPUT
    SEP : BYTE;
  END_VAR
  VAR_IN_OUT
    LIST : STRING[LIST_LENGTH];
  END_VAR
  VAR
    pt : PTR_TO OSCAT_BASIC_ARRAY1_LIST_LENGTH_OF_BYTE; // ARRAY[1..LIST_LENGTH] OF BYTE;
    read : INT := 1;
    write : INT := 1;
    last: BYTE;
    c: BYTE;
  END_VAR

  pt := ADR(LIST);

  FOR read := 1 TO LIST_LENGTH DO
    c := pt^[read];               (* read character from list *)
    IF c = 0 THEN EXIT;           (* exit the loop if character definbes end of string *)
    ELSIF (c <> SEP) OR (sep <> last) THEN  (* copy element from read to write position unless a double sep character is present *)
      pt^[write] := c;
      write := write + 1;
    END_IF;
    last := c;                  (* remember last character *)
  END_FOR;

  IF last = SEP THEN write := write - 1; END_IF;    (* if last character is sep then delete empty element at end *)
  IF write <= STRING_LENGTH THEN pt^[write] := 0;  END_IF;    (* terminate string with 0 *)

  LIST_CLEAN := TRUE;           (* retrun TRUE *)

(* revision histroy
  hm  28. jun. 2008 rev 1.0
    original release

  hm  19. jan. 2011 rev 1.1
    changed string(255) to string[LIST_LENGTH]

  hm  21. mar. 2011 rev 2.0
    all elements start with SEP
*)
END_FUNCTION

(* @PATH := '\/List Processing' *)
FUNCTION LIST_GET : STRING[LIST_LENGTH]
(*
  LIST_GET liefert das element an der stelle pos einer liste.
  die liste liegt als string von elementen vor die mit den zeichen SEP am anfang makiert sind.

  version 2.0 21. mar. 2011
  programmer  hugo
  tested by   oscat
*)
  VAR_INPUT
    SEP : BYTE;
    POS : INT;
  END_VAR
  VAR_IN_OUT
    LIST : STRING[LIST_LENGTH];
  END_VAR
  VAR
    i : INT := 1;
    o : INT := 1;
    pt : PTR_TO OSCAT_BASIC_ARRAY1_LIST_LENGTH_OF_BYTE; // ARRAY[1..LIST_LENGTH] OF BYTE;
    po : PTR_TO OSCAT_BASIC_ARRAY1_LIST_LENGTH_OF_BYTE; // ARRAY[1..LIST_LENGTH] OF BYTE;
    cnt: INT := 0;
    c: BYTE;
  END_VAR

  pt := ADR(LIST);              (* load pointers *)
//  po := ADR(LIST_GET);
  {asm}
    LEAX  __fc__LIST_GET
    WRX   po
  {end_asm}

  REPEAT
    c := pt^[i];
    IF cnt = pos THEN           (* copy element to output string *)
      IF c = SEP  THEN EXIT; END_IF;    (* next element stop copy and finish *)
      po^[o] := c;
      o := o + 1;
    ELSIF c = SEP THEN
      cnt := cnt + 1;
    END_IF;
    i := i + 1;
  UNTIL
    (i = LIST_LENGTH) OR (c = 0)
  END_REPEAT;
  po^[o] := 0;            (* close the output string *)

(* revision history
  hm  20. jun. 2008 rev 1.0
    original release

  hm  19. jan. 2011 rev 1.1
    changed string(255) to strring[LIST_LENGTH]

  hm  21. mar. 2011 rev 2.0
    all list elements start with SEP
*)
END_FUNCTION

(* @PATH := '\/List Processing' *)
FUNCTION LIST_INSERT : BOOL
(*
  LIST_INSERT setzt ein element an der stelle pos in eine liste ein.
  die liste liegt als string von elementen vor die mit den zeichen SEP am anfang markiert sind.

  version 2.0 21. mar. 2011
  programmer  hugo
  tested by   oscat
*)
  VAR_INPUT
    SEP : BYTE;
    POS : INT;
    INS : STRING[LIST_LENGTH];
  END_VAR
  VAR_IN_OUT
    LIST : STRING[LIST_LENGTH];
  END_VAR
  VAR
    pt : PTR_TO OSCAT_BASIC_ARRAY1_LIST_LENGTH_OF_BYTE; // ARRAY[1..LIST_LENGTH] OF BYTE;
    read : INT := 1;
    cnt : INT := 1;
    sx : STRING[1];
  END_VAR

  (* load pointers *)
  pt := ADR(LIST);

  IF LEN(ins) + 1 + LEN(LIST) > LIST_LENGTH THEN
    LIST_INSERT := FALSE;
  ELSE
    LIST_INSERT := TRUE;
    (* search for position *)
    WHILE read < LIST_LENGTH DO
      IF cnt >= POS THEN
        sx := CHR_TO_STRING(SEP);
        INS := CONCAT(sx, INS);
        LIST := INSERT(LIST, INS, read - 1);
        LIST_INSERT := TRUE;
        RETURN;
      END_IF;
      IF pt^[read]  = 0 THEN        (* list is too short add empty element *)
        pt^[read] := SEP;
        pt^[read + 1] := 0;
      END_IF;
      read := read + 1;
      IF (pt^[read] = SEP) OR (pt^[read] = 0) THEN cnt := cnt + 1; END_IF;
    END_WHILE;
  END_IF;

(* revision history
  hm  28. jun. 2008 rev 1.0
    original release

  hm  17. dec. 2008 rev 1.1
    changes name of function chr to chr_to_string

  hm  19. jan. 2011 rev 1.2
    changed string(255) to string[LIST_LENGTH]

  hm  21. mar. 2011 rev 2.0
    all list elements start with SEP
*)
END_FUNCTION

(* @PATH := '\/List Processing' *)
FUNCTION LIST_LEN : INT
(*
  LIST_LEN liefert die anzahl der elemente einer liste.
  die liste liegt als string von elementen vor die mit den zeichen SEP am anfang markiert sind.

  version 2.0 21. mar. 2011
  programmer  hugo
  tested by   oscat
*)
  VAR_INPUT
    SEP : BYTE;
  END_VAR
  VAR_IN_OUT
    LIST : STRING[LIST_LENGTH];
  END_VAR
  VAR
    pt : PTR_TO OSCAT_BASIC_ARRAY1_LIST_LENGTH_OF_BYTE; // ARRAY[1..LIST_LENGTH] OF BYTE;
    pos: INT := 1;
    c: BYTE;
  END_VAR

  pt := ADR(LIST);
  LIST_LEN := 0;
  REPEAT
  	c := pt^[pos];
  	IF c = SEP THEN LIST_LEN := LIST_LEN + 1; END_IF;
  	pos := pos + 1;
  UNTIL
  	(c = 0) OR (pos > LIST_LENGTH)
  END_REPEAT;

(* revision history
  hm  25. jun. 2008 rev 1.0
    original release

  hm  16. oct. 2008 rev 1.1
    fixed a problem where list_len would only work up to LIST_LENGTH

  hm  19. jan. 2001 rev 1.2
    changed string(255) to string[LIST_LENGTH]

  hm  21. mar. 2011 rev 2.0
    all list elements start with SEP
*)
END_FUNCTION

(* @PATH := '\/List Processing' *)
FUNCTION_BLOCK LIST_NEXT
(*
  LIST_NEXT retrieves the next element of a list, starting from element 1 after reset or first init.
  when the end of the lisat is reached a '' empty string is returned and NUL is set to true.
  die liste liegt als string von elementen vor die mit den zeichen SEP am anfang markiert sind.

  version 2.0 21. mar. 2011
  programmer  hugo
  tested by   oscat
*)
  VAR_INPUT
    SEP : BYTE;
    RST : BOOL;
  END_VAR
  VAR_IN_OUT
    LIST : STRING[LIST_LENGTH];
  END_VAR
  VAR_OUTPUT
    LEL : STRING[LIST_LENGTH];
    NUL : BOOL;
  END_VAR
  VAR
    pos : INT := 1;
    pt : PTR_TO OSCAT_BASIC_ARRAY1_LIST_LENGTH_OF_BYTE; // ARRAY[1..LIST_LENGTH] OF BYTE;
    po : PTR_TO OSCAT_BASIC_ARRAY1_LIST_LENGTH_OF_BYTE; // ARRAY[1..LIST_LENGTH] OF BYTE;
    c: BYTE;
    write: INT;
  END_VAR

  pt := ADR(LIST);
  po := ADR(LEL);

  IF rst THEN
    pos := 1;
  END_IF;

  IF (pt^[pos] = 0) OR (pos = LIST_LENGTH) THEN
    LEL := '';
    NUL := TRUE;
  ELSE
    NUL := FALSE;
    write := 1;
    FOR pos := pos + 1 TO LIST_LENGTH DO
      c := pt^[pos];
      IF (c = 0) OR (c = SEP) THEN
        po^[write] := 0;
        RETURN;
      ELSE
        po^[write] := pt^[pos];
        write := write + 1;
      END_IF;
    END_FOR;
  END_IF;

(* revision history
  hm  25. jun. 2008 rev 1.0
    original release

  hm  19. jan. 2011 rev 1.1
    changed string(255) to string[LIST_LENGTH]

  hm  21. mar. 2011 rev 2.0
    all elements start with SEP
*)
END_FUNCTION_BLOCK

(* @PATH := '\/List Processing' *)
FUNCTION LIST_RETRIEVE : STRING[LIST_LENGTH]
(*
  LIST_RETRIEVE liefert das element an der stelle pos einer liste und löscht das element aus der liste.
  die liste liegt als string von elementen vor die mit den zeichen SEP separiert sind.

  version 2.0   21. mar. 2011
  programmer  hugo
  tested by   oscat
*)
  VAR_INPUT
    SEP : BYTE;
    POS : INT;
  END_VAR
  VAR_IN_OUT
    LIST : STRING[LIST_LENGTH];
  END_VAR
  VAR
    i : INT;
    o : INT := 1;
    w : INT := 1;
    pt : PTR_TO OSCAT_BASIC_ARRAY1_LIST_LENGTH_OF_BYTE; // ARRAY[1..LIST_LENGTH] OF BYTE;
    po : PTR_TO OSCAT_BASIC_ARRAY1_LIST_LENGTH_OF_BYTE; // ARRAY[1..LIST_LENGTH] OF BYTE;
    cnt: INT := 0;
    c: BYTE;
  END_VAR

  (* load pointers *)
  pt := ADR(LIST);
//  po := ADR(LIST_RETRIEVE);
  {asm}
    LEAX  __fc__LIST_RETRIEVE
    WRX   po
  {end_asm}

  IF pos > 0 THEN
    FOR i := 1 TO LIST_LENGTH DO
      c := pt^[i];
      IF c = 0 THEN
        po^[o] := 0;
        IF cnt < pos THEN pt^[w + 1] := 0; ELSE pt^[w] := 0; END_IF;
        RETURN;
      ELSIF cnt = pos AND c <> SEP THEN       (* we have found the element *)
        po^[o] := pt^[i];
        o := o + 1;
      ELSIF cnt >= pos THEN
        pt^[w] := c;
        w := w + 1;
      ELSE
        w := i;
      END_IF;
      IF c = sep THEN cnt := cnt + 1; END_IF;
    END_FOR;
  ELSE
    LIST_RETRIEVE := '';
  END_IF;

(* revision history
  hm  28. jun. 2008 rev 1.0
    original release

  hm  19. jan. 2011 rev 1.1
    changed string(255) to string[LIST_LENGTH]

  hm  21. mar. 2011 rev 2.0
    all elements start with SEP
*)
END_FUNCTION

(* @PATH := '\/List Processing' *)
FUNCTION LIST_RETRIEVE_LAST : STRING[LIST_LENGTH]
(*
  LIST_RETRIEVE_LAST liefert das letzte element einer liste und löscht das element aus der liste.
  die liste liegt als string von elementen vor die mit den zeichen SEP beginnen.

  version 2.0   21. mar. 2011
  programmer  hugo
  tested by   oscat
*)
  VAR_INPUT
    SEP : BYTE;
  END_VAR
  VAR_IN_OUT
    LIST : STRING[LIST_LENGTH];
  END_VAR
  VAR
    i : INT;
    last : INT := 1;
    pt : PTR_TO OSCAT_BASIC_ARRAY1_LIST_LENGTH_OF_BYTE; // ARRAY[1..LIST_LENGTH] OF BYTE;
    c: BYTE;
  END_VAR

  (* load pointers *)
  pt := ADR(LIST);

  (* search position of last element *)
  FOR i := 1 TO LIST_LENGTH DO
    c := pt^[i];
    IF c = 0 THEN
      EXIT;
    ELSIF C = SEP THEN
      last := i;
    END_IF;
  END_FOR;
  (* return last element of list *)
  LIST_RETRIEVE_LAST := MID(LIST, LIST_LENGTH, last + 1);
  (* terminate list at i *)
  pt^[last] := 0;

(* revision history
  hm  21. mar. 2011 rev 2.0
    new module
*)
END_FUNCTION

(* ---- OscatBasicLib_333a.st ---- *)
VAR_GLOBAL CONSTANT
	STRING_LENGTH : INT := 250;
	LIST_LENGTH : INT := 250;
END_VAR

(* revision history
  hm 3. mar. 2007
  	extended accuracy of pi2
  	renamed T0 to Tk for better compatibility with other libraries
  	renamed C t0 c0 for better compatibility

  hm	2. may. 2007
  	added RU universal gas constant

  hm	1. oct. 2007
  	added setup parameter STEP7

  hm 31. oct. 2007
  	added PN

  hm	6. mar. 2008
  	added setup Parameter EXTENDED_ASCII

  hm	28. Mar. 2008
  	added setup parameter STRING_LENGTH

  hm	7. apr. 2008
  	Deleted unused setup parameter Step7

  hm	19. apr. 2008
  	added setup parameter NETWORK_BUFFER_SIZE

  hm	27. apr. 2008
  	added PI05 and PI025

  hm	18. may. 2008
  	added charname lists
  	renamed E to E1

  hm	30. jun. 2008
  	reduced size of string constants to 253 to avoid problems with target aixia DCUF

  hm	21. sep. 2008
  	added section language setup
  	added section location setup

  hm	20. oct. 2008
  	changed to structured constants

  hm	16. nov. 2008
  	moved structured constants to global vars for compatibility reasons

  hm	13. nov. 2009
  	added network_buffer_short_size
  	renamed network_buffer_long_size
  	changed string length to 250

  hm	20. jan. 2011
  	removed network buffers
  	added list_length
*)

TYPE CONSTANTS_SETUP :
  STRUCT
    (* setup Parameters *)
    EXTENDED_ASCII : BOOL := TRUE;                  (* extends the ASCII character set to special characters eg ÄÖÜ *)
    CHARNAMES : ARRAY[1..4] OF STRING[253] := [     (* stores Unicode character names *)
      ';"&quot;&&amp;<&lt;>&gt;€&euro; &nbsp;?&iexcl;?&cent;L&pound;¤&curren;A&yen;¦&brvbar;§&sect;¨&uml;©&copy;S&ordf;«&laquo;¬&not;­&shy;®&reg;Z&macr;°&deg;±&plusmn;?&sup2;l&sup3;´&acute;µ&micro;¶&para;·&middot;¸&cedil;a&sup1;s&ordm;»&raquo;L&frac14;U&Ucirc;',
      ';l&frac34;z&iquest;R&Agrave;Á&Aacute;Â&Acirc;A&Atilde;Ä&Auml;L&Aring;C&AElig;Ç&Ccedil;C&Egrave;É&Eacute;E&Ecirc;Ë&Euml;E&Igrave;Í&Iacute;Î&Icirc;D&Iuml;Ð&ETH;N&Ntilde;N&Ograve;Ó&Oacute;Ô&Ocirc;O&Otilde;Ö&Ouml;×&times;R&Oslash;U&Ugrave;Ú&Uacute;?&frac12;',
      ';Ü&Uuml;Ý&Yacute;T&THORN;ß&szlig;r&agrave;á&aacute;â&acirc;a&atilde;ä&auml;l&aring;c&aelig;ç&ccedil;c&egrave;é&eacute;e&ecirc;ë&euml;e&igrave;í&iacute;î&icirc;d&iuml;d&eth;n&ntilde;n&ograve;ó&oacute;ô&ocirc;o&otilde;ö&ouml;÷&divide;r&oslash;u&ugrave;',
      ';ú&uacute;u&ucirc;ü&uuml;ý&yacute;t&thorn;?&yuml;'];
    MTH_OFS : ARRAY[1..12] OF INT := [0,31,59,90,120,151,181,212,243,273,304,334];
    DECADES : ARRAY[0..8] OF REAL := [1.0,10.0,100.0,1000.0,10000.0,10000.0,100000.0,1000000.0,10000000.0];
  END_STRUCT;
END_TYPE

(* revision history
  hm  24.10.2008  rev 1.0
    original version
*)

TYPE CONSTANTS_MATH :
  STRUCT
    PI : REAL :=  3.14159265358979323846; //???3.14159265358979323846264338327950288;    (* Kreiszahl PI *)
    PI2 : REAL :=   6.28318530717958647692;//???6.28318530717958647692528676655900576;  (* PI * 2 *)
    PI4 : REAL :=  12.56637061435917295385;//???12.56637061435917295385057353311801152;  (* PI * 4 *)
    PI05 : REAL :=  1.5707963267949;              (* PI / 2 *)
    PI025 : REAL := 0.785398163397448;              (* PI / 4 *)
    PI_INV : REAL := 0.318309886183791;           (* 1 / PI *)
    E : REAL :=   2.71828182845904523536;//???2.71828182845904523536028747135266249;    (* Euler constant e *)
    E_INV : REAL := 0.367879441171442;              (* 1 / e *)
    SQ2 : REAL := 1.4142135623731;              (* Root of 2 *)
    FACTS : ARRAY[0..12] OF DINT := [1,1,2,6,24,120,720,5040,40320,362880,3628800,39916800,479001600]; (* Faculties 0-12 *)
  END_STRUCT;
END_TYPE

(* revision history
  hm  26.10.2008  rev 1.0
    original version

  hm  26. mar. 2011 rev 1.1
    added array facts
*)

TYPE FRACTION :
  STRUCT
    NUMERATOR : INT;     (* Numerator of the fraction *)
    DENOMINATOR : INT;   (* Denominator of the fraction *)
  END_STRUCT;
END_TYPE

TYPE REAL2 :
  STRUCT
    R1 : REAL;  (* small value *)
    RX : REAL;  (* big value *)
  END_STRUCT;
END_TYPE

(* revision history
  hm  18. oct. 2008
    original version
*)

TYPE SDT :             (* defnes a structured time-date format *)
  STRUCT
    YEAR : INT;
    MONTH : INT;
    DAY : INT;
    WEEKDAY : INT;
    HOUR : INT;
    MINUTE : INT;
    SECOND : INT;
    MS : INT;
  END_STRUCT;
END_TYPE

(* revision history
  hm  18. oct. 2008
    original version
*)

TYPE TIMER_EVENT :
  STRUCT
    TYP : BYTE;            (* Event Type *)
    CHANNEL : BYTE;        (* Channel *)
    DAY : BYTE;            (* Day or days *)
    START : TOD;           (* Start time *)
    DURATION : TIME;       (* Duration *)
    LAND : BYTE;           (* Logical AND *)
    LOR : BYTE;            (* Logical OR *)
    LAST : DT;             (* last activity of the event *)
  END_STRUCT;
END_TYPE

(* revision history
hm  18. oct. 2008 rev 1.0
  original version

hm  26. jan. 2011 rev 1.1
  changed type of last to be DT
*)

TYPE CALENDAR :
  STRUCT
    UTC : DT;            (* world time UTC *)
    LDT : DT;            (* local time *)
    LDATE : DATE;        (* local date *)
    LTOD : TOD;          (* local time of day *)
    YEAR : INT;          (* year of LDATE *)
    MONTH : INT;         (* month of LDATE *)
    DAY : INT;           (* day of LDATE *)
    WEEKDAY : INT;       (* weekday of LDATE *)
    OFFSET : INT;        (* Time Zone Offset for Local time in minutes *)
    DST_EN : BOOL;       (* daylight savings time enable *)
    DST_ON : BOOL;       (* true when daylight savings time os on *)
    NAME : STRING[5];    (* name of time zone *)
    LANGUAGE : INT;      (* location number pls see location setup *)
    LONGITUDE : REAL;    (* longitude of current location *)
    LATITUDE : REAL;     (* latitude of current location *)
    SUN_RISE : TOD;      (* sun_rise for current location *)
    SUN_SET : TOD;       (* sun_set for current location *)
    SUN_MIDDAY : TOD;    (* worldtime when sun stands at south position *)
    SUN_HEIGTH : REAL ;  (* suns heigth at midday, south position *)
    SUN_HOR : REAL;      (* sun angle horizontal 0 = north in degrees *)
    SUN_VER : REAL;      (* sun angle vertical above horizon in degrees *)
    NIGHT : BOOL;        (* true between sun_set and sun_rise *)
    HOLIDAY : BOOL;      (* true when holiday *)
    HOLY_NAME : STRING[30]; (* name of holiday *)
    WORK_WEEK : INT;      (* current work week *)
  END_STRUCT;
END_TYPE

(* revision history
  hm  21. nov. 2008 rev 1.0
    original version

  hm  8. feb. 2009  rev 1.1
    added sun position data

  hm  10. mar. 2009 rev 1.2
    added work_week, sun_midday, sun_heigth

  hm  23. jan 2010  rev 1.3
    sun_rise, sun_set and sun_midday are now calculated in local time
*)

TYPE ESR_DATA :                 (* ESR_DATA is used for Error and Status Reporting modules *)
  STRUCT
    TYP : BYTE;                 (* Data Type *)
    ADRESS : STRING[10];        (* Adress designation *)
    DS : DT;                    (* Date / time stamp *)
    TS : TIME;                  (* Timestamp in milliseconds *)
    DATA : ARRAY[0..7] OF BYTE; (* Data packet *)
  END_STRUCT;
END_TYPE

(* revision history
  hm  18. oct. 2008
    original version
*)

TYPE HOLIDAY_DATA :
  STRUCT
    NAME : STRING[30];      (* Name of the holiday *)
    DAY : SINT;             (* Day of public holiday *)
    MONTH : SINT;           (* Month of the holy day *)
    USE : SINT;             (* activates the holyday (0=off, 1=on) *)
  END_STRUCT;
END_TYPE

(* revision history
  hm  18. oct. 2008
    original version
*)
(* if month = 0 then F_day is the offset in days from easter
   used :0 = NOT used, 1 = used, -1..-7 menas the weekday before the specified DATE example -3 means wednesday before 23.11
*)
(* samples for Holiday data

  HOLIDAY_DE : ARRAY[0..29] OF HOLIDAY_DATA := (name := 'Neujahr', day := 1, month := 1, use := 1),
    (name := 'Heilig Drei Könige', day := 6, month := 1, use := 1),
    (name := 'Karfreitag', day := -2, month := 0, use := 1),
    (name := 'Ostersonntag', day := 0, month := 0, use := 1),
    (name := 'Ostermontag', day := 1, month := 0, use := 1),
    (name := 'Tag der Arbeit', day := 1, month := 5, use := 1),
    (name := 'Christi Himmelfahrt', day := 39, month := 0, use := 1),
    (name := 'Pfingstsonntag', day := 49, month := 0, use := 1),
    (name := 'Pfingstmontag', day := 50, month := 0, use := 1),
    (name := 'Fronleichnam', day := 60, month := 0, use := 1),
    (name := 'Augsburger Friedensfest', day := 8, month := 8, use := 0),
    (name := 'Maria Himmelfahrt', day := 15, month := 8, use := 1),
    (name := 'Tag der Deutschen Einheit', day := 3, month := 10, use := 1),
    (name := 'Reformationstag', day := 31, month := 10, use := 0),
    (name := 'Allerheiligen', day := 1, month := 11, use := 1),
    (name := 'Buss und Bettag', day := 23, month := 11, use := 0),
    (name := '1. Weihnachtstag', day := 25, month := 12, use := 1),
    (name := '2. Weihnachtstag', day := 26, month := 12, use := 1);

  HOLIDAY_AT : ARRAY[0..29] OF HOLIDAY_DATA := (name := 'Neujahr', day := 1, month := 1, use := 1),
    (name := 'Heilig Drei Könige', day := 6, month := 1, use := 1),
    (name := 'Karfreitag', day := -2, month := 0, use := 1),
    (name := 'Ostersonntag', day := 0, month := 0, use := 1),
    (name := 'Ostermontag', day := 1, month := 0, use := 1),
    (name := '', day := 1, month := 5, use := 0),
    (name := 'Christi Himmelfahrt', day := 39, month := 0, use := 1),
    (name := 'Pfingstsonntag', day := 49, month := 0, use := 1),
    (name := 'Pfingstmontag', day := 50, month := 0, use := 1),
    (name := 'Fronleichnam', day := 60, month := 0, use := 1),
    (name := '', day := 8, month := 8, use := 0),
    (name := 'Maria Himmelfahrt', day := 15, month := 8, use := 1),
    (name := '', day := 3, month := 10, use := 0),
    (name := '', day := 31, month := 10, use := 0),
    (name := 'Allerheiligen', day := 1, month := 11, use := 1),
    (name := 'Maria Empfängnis', day := 8, month := 12, use := 1),
    (name := '1. Weihnachtstag', day := 25, month := 12, use := 1),
    (name := '2. Weihnachtstag', day := 26, month := 12, use := 1);

  HOLIDAY_FR : ARRAY[0..29] OF HOLIDAY_DATA := (name := 'Nouvel an', day := 1, month := 1, use := 1),
    (name := 'St Valentin', day := 14, month := 2, use := 0),
    (name := 'Vendredi Saint (alsace)', day := -2, month := 0, use := 0),
    (name := 'Dimanche de pâques', day := 0, month := 0, use := 1),
    (name := 'Lundi de pâques', day := 1, month := 0, use := 1),
    (name := 'Jeudi de Ascension', day := 39, month := 0, use := 1),
    (name := 'dimanche de Pentecôte ', day := 49, month := 0, use := 1),
    (name := 'jeudi de la Trinité', day := 60, month := 0, use := 0),
    (name := 'Fete du travail', day := 1, month := 5, use := 1),
    (name := 'Victoire 1945 ', day := 8, month := 5, use := 1),
    (name := 'Prise de La bastille', day := 14, month := 7, use := 1),
    (name := '15 Aout 1944', day := 15, month := 8, use := 1),
    (name := 'Halloween', day := 31, month := 10, use := 0),
    (name := 'Armistice 1918', day := 11, month := 11, use := 1),
    (name := 'Noël', day := 25, month := 12, use := 1),
    (name := 'Saint Étienne (alsace)', day := 26, month := 12, use := 0),
    (name := 'Fete de la musique', day := 21, month := 6, use := 0);

  HOLIDAY_BED : ARRAY[0..29] OF HOLIDAY_DATA := (name := 'Neujahr', day := 1, month := 1, use := 1),
    (name := 'Ostersonntag', day := 0, month := 0, use := 1),
    (name := 'Ostermontag', day := 1, month := 0, use := 1),
    (name := 'Tag der Arbeit', day := 1, month := 5, use := 1),
    (name := 'Christi Himmelfahrt', day := 39, month := 0, use := 1),
    (name := 'Pfingsten', day := 49, month := 0, use := 1),
    (name := 'Pfingstmontag', day := 50, month := 0, use := 1),
    (name := 'Nationalfeiertag', day := 21, month := 7, use := 1),
    (name := 'Mariä Himmelfahrt', day := 15, month := 8, use := 1),
    (name := 'Allerheiligen', day := 1, month := 11, use := 1),
    (name := 'Feiertag DG', day := 15, month := 11, use := 1),
    (name := 'Heiligabend', day := 24, month := 12, use := 1),
    (name := '1. Weihnachtstag', day := 25, month := 12, use := 1),
    (name := '2. Weihnachtstag', day := 26, month := 12, use := 1),
    (name := 'Silvester', day := 31, month := 12, use := 1);

  HOLIDAY_ITD : ARRAY[0..29] OF HOLIDAY_DATA := (name := 'Neujahr', day := 1, month := 1, use := 1),
    (name := 'Heilig Drei Könige', day := 6, month := 1, use := 1),
    (name := 'Ostersonntag', day := 0, month := 0, use := 1),
    (name := 'Ostermontag', day := 1, month := 0, use := 1),
    (name := 'Tag der Befeiung Italiens', day := 25, month := 4, use := 1),
    (name := 'Tag der Arbeit', day := 1, month := 5, use := 1),
    (name := 'Pfingsten', day := 49, month := 0, use := 1),
    (name := 'Pfingstmontag', day := 50, month := 0, use := 1),
    (name := 'Tag der Republik Italien', day := 2, month := 6, use := 1),
    (name := 'Mariä Himmelfahrt', day := 15, month := 8, use := 1),
    (name := 'Allerheiligen', day := 1, month := 11, use := 1),
    (name := 'Mariä Empfängnis', day := 8, month := 12, use := 1),
    (name := 'Heiligabend', day := 24, month := 12, use := 0),
    (name := '1. Weihnachtstag', day := 25, month := 12, use := 1),
    (name := '2. Stephanstag', day := 26, month := 12, use := 1);
*)

TYPE COMPLEX :   (* structure can present complex numbers *)
  STRUCT
    re : REAL;   (*Real part of a complex number*)
    im : REAL;   (*Imaginary part of a complex number*)
  END_STRUCT;
END_TYPE

(* revision history
  hm  18. oct. 2008
    original version
*)

TYPE VECTOR_3 :   (* stores the three vectors of a three-dimensional vector space *)
  STRUCT
    X : REAL;
    Y : REAL;
    Z : REAL;
  END_STRUCT;
END_TYPE

(* revision history
  hm  18. oct. 2008
    original version
*)

TYPE CONSTANTS_LANGUAGE :
  STRUCT
    (* Language Setup *)
    DEFAULT : INT := 1; (* 1=english, 2=german 3=french *)
    LMAX    : INT := 3; (* specifes how many languages are available *)
    WEEKDAYS : ARRAY[1..3, 1..7] OF STRING[10] := [
                            'Monday', 'Tuesday', 'Wednesday', 'Thursday', 'Friday', 'Saturday', 'Sunday',
                            'Montag', 'Dienstag', 'Mittwoch', 'Donnerstag', 'Freitag', 'Samstag', 'Sonntag',
                            'Lundi', 'Mardi', 'Mercredi', 'Jeudi', 'Vendredi', 'Samedi', 'Dimanche'];
    WEEKDAYS2 : ARRAY[1..3, 1..7] OF STRING[2] := [
                            'Mo', 'Tu', 'We', 'Th', 'Fr', 'Sa', 'Su',
                            'Mo', 'Di', 'Mi', 'Do', 'Fr', 'Sa', 'So',
                            'Lu', 'Ma', 'Me', 'Je', 'Ve', 'Sa', 'Di'];
    MONTHS : ARRAY[1..3, 1..12] OF STRING[10] := [
                            'January', 'February', 'March', 'April', 'May', 'June', 'July', 'August', 'September', 'October', 'November', 'December',
                            'Januar', 'Februar', 'März', 'April', 'Mai', 'Juni', 'Juli', 'August', 'September', 'Oktober', 'November', 'Dezember',
                            'Janvier', 'Février', 'mars', 'Avril', 'Mai', 'Juin', 'Juillet', 'Aout', 'Septembre', 'Octobre', 'Novembre', 'Decembre'];
    MONTHS3 : ARRAY[1..3, 1..12] OF STRING[3] := [
                            'Jan', 'Feb', 'Mar', 'Apr', 'May', 'Jun', 'Jul', 'Aug', 'Sep', 'Oct', 'Nov', 'Dec',
                            'Jan', 'Feb', 'Mrz', 'Apr', 'Mai', 'Jun', 'Jul', 'Aug', 'Sep', 'Okt', 'Nov', 'Dez',
                            'Jan', 'Fev', 'Mar', 'Avr', 'Mai', 'Jun', 'Jul', 'Aou', 'Sep', 'Oct', 'Nov', 'Dec'];
    DIRS : ARRAY[1..3,0..15] OF STRING[3] := [
                            'N', 'NNE', 'NE', 'ENE', 'E', 'ESE', 'SE', 'SSE', 'S', 'SSW', 'SW', 'WSW', 'W', 'WNW', 'NW', 'NNW',
                            'N', 'NNO', 'NO', 'ONO', 'O', 'OSO', 'SO', 'SSO', 'S', 'SSW', 'SW', 'WSW', 'W', 'WNW', 'NW', 'NNW',
                            'N', 'NNO', 'NO', 'ONO', 'O', 'OSO', 'SO', 'SSO', 'S', 'SSW', 'SW', 'WSW', 'W', 'WNW', 'NW', 'NNW'];
  END_STRUCT;
END_TYPE

(* revision history
  hm  19. oct. 2008 rev 1.0
    original version

  hm  22. oct. 2008 rev 1.1
    added directions DIRS

  hm  23. dec. 2008 rev 1.2
    added french language
*)

TYPE CONSTANTS_LOCATION :
  STRUCT
    (* location setup *)
    DEFAULT : INT := 1;                                (* 1=germany, 2=austria 3=france 4=belgium-german 5= italien-Südtirol *)
    LMAX : INT := 5;                                   (* indicates how many places are defned *)
    LANGUAGE : ARRAY[1..5] OF INT := [ 2, 2, 3, 2, 2]; (* language spoken in the location *)
  END_STRUCT;
END_TYPE

(* revision history
  hm  20. oct. 2008 rev 1.0
    original version

  hm  23. dec. 2008 rev 1.1
    added french holidays

  hm  18. jan 2011  rev 1.2
    added spoken language
    deleted holidays from structure for more flexibility
*)

TYPE CONSTANTS_PHYS :
  STRUCT
    C : REAL := 299792458.0;        (* Lichtgeschwindigkeit in m/s *)
    E : REAL := 1.60217653E-19;     (* elementarladung in Colomb = A * s *)
    G : REAL := 9.80665;            (* Erdbeschleunigung in m / s? *)
    T0 : REAL := -273.15;           (* absoluter Nullpunkt in °C *)
    RU : REAL := 8.314472;          (* Universelle Gaskonstante in J / (mol · K) *)
    PN : REAL := 101325.0;          (* NormalDruck in Pa *)
  END_STRUCT;
END_TYPE

(* revision history
  hm  18.10.2008  rev 1.0
    original version

  hm  13. mar. 2009 rev 1.1
    real constants updated to new systax using dot
*)

VAR_GLOBAL
  MATH     : CONSTANTS_MATH;
  PHYS     : CONSTANTS_PHYS;
  LANGUAGE : CONSTANTS_LANGUAGE;
  SETUP    : CONSTANTS_SETUP;
  LOCATION : CONSTANTS_LOCATION;
END_VAR
